Fanuc KAREL source: KD00046.KL

PROGRAM KD00046
%NOLOCKGROUP
%DEFGROUP = 1
VAR
  I: INTEGER
  J: INTEGER
  B: BOOLEAN
  R: REAL
  S: STRING[80]
  V: VECTOR
BEGIN
  V.X = 1.0
  MOVE RELATIVE V
END KD00046
